(* IEC 61131-3 sources: openplc-runtime/tests/hmi_e2e/project/pous/programs, 1 file *)

(* ---- Main.st ---- *)
PROGRAM Main
  VAR
    Run : BOOL;
    Level : REAL;
    Setpoint : INT;
  END_VAR

  IF Run THEN
    Level := Level + 1.0;
  END_IF;
END_PROGRAM
